Fanuc KAREL source: KC00001.KL

PROGRAM KC00001
%NOLOCKGROUP
%ENVIRONMENT PC
VAR
  I: INTEGER
  J: INTEGER
  K: INTEGER
  R: REAL
  B: BOOLEAN
  S: STRING[80]
  T: STRING[80]
  P: PATH
  Q: PATH
  AI: ARRAY[8] OF INTEGER
  AB: ARRAY[244] OF BYTE
BEGIN
  S = 'P'
  T = 'I'
  ADD_BYNAMEPC(AB,I,S,T,J)
END KC00001
